Fanuc KAREL source: KT00739.KL

PROGRAM KT00739
%NOLOCKGROUP
VAR
  ARG: ARRAY[4] OF BYTE
  OUT: INTEGER
BEGIN
  OUT = ARRAY_LEN(ARG)
END KT00739
